Fanuc KAREL source: kx00006.KL

-- PROVISIONAL review KL for V940-1; original PC SHA256 6e68b6597779d4205dfaf2d55d34cf3394302bb21e014c91ea62e1c90404ac3c
-- Incomplete behavior may be omitted. Consult companion uncertainty JSON. Do not deploy.
PROGRAM KX00006
%NOLOCKGROUP
VAR
  I : INTEGER
  J : INTEGER
  B : BOOLEAN
  F : FILE
  S : STRING[80]
-- UNRESOLVED_DECL P type=000102
BEGIN
  -- V9_ZERO_TABLE_METADATA_HINT layout=0001; no indexed target words; source/name/runtime held
  -- UNRESOLVED_PC offsets 5-13; opcodes 9D,2E,0F
  -- UNRESOLVED_PC offsets 18-22; opcodes 7F
END KX00006
